(* IEC 61131-3 sources: plc-iiot-stack/src/POUs/Iiot/FB_MqttDiag, 14 files *)

(* ---- FB_MqttDiag.decl.st ---- *)
// Назначение: ведение связи с брокером и состояние узла (data_schema 6): автомат Disabled -> Connecting ->
//             Connected -> Backoff -> Connecting; тайм-аут подключения, пауза между попытками удваивается от
//             tBackoffMin до tBackoffMax и снова минимальна после tStable устойчивой связи. Перед Connect —
//             завещание (LWT) в <prefix>/<sNode>/status/connection: offline/lwt со временем подключения;
//             после подключения — рождение online/birth (source, sw_version, period_ms), затем xReady.
//             Выключение при связи — offline/shutdown, разрыв в следующем вызове. Без часов ПЛК обмен не
//             начинается (MQTT_ERR_NO_CLOCK). Счётчики, код последней ошибки, сводный статус в духе NE 107.
// Автор:      kr0nsch
// Версия:     0.1.0
// Документ:   docs/plc_mqtt.md, раздел «Связь и состояние узла»
FUNCTION_BLOCK FB_MqttDiag
VAR_INPUT
    xEnable : BOOL;
    itfClient : I_MqttClient;
    ltNow : LTIME;                                            // монотонное время (LTIME())
    uliTs_ms : ULINT;                                         // время UTC, мс (поле ts)
    sTopicPrefix : STRING(GVL_Const.IIOT_PREFIX_LEN);         // site/area/unit
    sNode : STRING(GVL_Const.IIOT_DEVICE_LEN) := 'PLC1';
    sSwVersion : STRING(GVL_Const.IIOT_TEXT_LEN) := '0.1.0';
    tPeriod : TIME := GVL_Const.TELEMETRY_PERIOD_DEFAULT;    // период контрольной публикации (period_ms)
    tConnectTimeout : TIME := GVL_Const.CONNECT_TIMEOUT_DEFAULT;
    tBackoffMin : TIME := GVL_Const.BACKOFF_MIN_DEFAULT;
    tBackoffMax : TIME := GVL_Const.BACKOFF_MAX_DEFAULT;
    tStable : TIME := GVL_Const.STABLE_TIME_DEFAULT;
    tDegradeWindow : TIME := GVL_Const.TELEMETRY_PERIOD_DEFAULT;   // окно оценки отказов публикаций
    uiFailThreshold : UINT := GVL_Const.FAIL_THRESHOLD_DEFAULT;
    udiPubFailed : UDINT;                                     // отказы публикаций телеметрии и тревог
END_VAR
VAR_IN_OUT
    stBroker : ST_MqttBrokerCfg;                              // ФБ дописывает топик и текст LWT
END_VAR
VAR_OUTPUT
    eState : E_MqttConnState := E_MqttConnState.Disabled;
    eNe107 : E_IiotNe107 := E_IiotNe107.CheckFunction;
    xConnected : BOOL;
    xReady : BOOL;                  // связь есть и рождение опубликовано: можно публиковать
    udiConnects : UDINT;            // успешных подключений
    udiDisconnects : UDINT;         // потерь установленной связи
    udiConnectFailures : UDINT;     // неудачных попыток подключения
    uiConsecutiveFailures : UINT;   // неудачных попыток подряд (сброс после tStable связи)
    diLastError : DINT;             // GVL_Const.MQTT_ERR_* или код библиотеки
    tBackoff : TIME;                // пауза перед следующей попыткой
    xDegraded : BOOL;               // за последнее окно публикации отклонялись
END_VAR
VAR
    ltStateSince : LTIME;
    ltDegradeStart : LTIME;
    udiPubFailedRef : UDINT;
    fbJson : FB_JsonBuilder;
    sTopic : STRING(GVL_Const.MQTT_TOPIC_LEN);
END_VAR

(* ---- BuildStatus.method.decl.st ---- *)
// JSON состояния узла в fbJson: online/birth (с source, sw_version, period_ms) или offline/<sReason>.
METHOD PRIVATE BuildStatus : BOOL
VAR_INPUT
    xOnline : BOOL;
    sReason : STRING(GVL_Const.IIOT_TEXT_LEN);
END_VAR

(* ---- BuildStatus.method.impl.st ---- *)
fbJson.Begin();
fbJson.AddString(sKey := 'schema_version', sValue := GVL_Const.IIOT_SCHEMA_VERSION);
fbJson.AddInt(sKey := 'ts', liValue := ULINT_TO_LINT(uliTs_ms));
fbJson.AddString(sKey := 'node', sValue := sNode);
IF xOnline THEN
    fbJson.AddString(sKey := 'state', sValue := 'online');
ELSE
    fbJson.AddString(sKey := 'state', sValue := 'offline');
END_IF
fbJson.AddString(sKey := 'reason', sValue := sReason);
IF xOnline THEN
    fbJson.AddString(sKey := 'source', sValue := GVL_Const.IIOT_SOURCE);
    fbJson.AddString(sKey := 'sw_version', sValue := sSwVersion);
    fbJson.AddInt(sKey := 'period_ms', liValue := ULINT_TO_LINT(TIME_TO_ULINT(tPeriod)));
END_IF
BuildStatus := fbJson.Finish();

(* ---- ConnectFailed.method.decl.st ---- *)
// Неудачная попытка подключения: код ошибки (клиента или diDefaultError), счётчики, разрыв, пауза.
METHOD PRIVATE ConnectFailed
VAR_INPUT
    diDefaultError : DINT;
END_VAR

(* ---- ConnectFailed.method.impl.st ---- *)
diLastError := itfClient.LastError();
IF diLastError = GVL_Const.MQTT_ERR_NONE THEN
    diLastError := diDefaultError;
END_IF
udiConnectFailures := udiConnectFailures + 1;
IF uiConsecutiveFailures < UINT#65535 THEN
    uiConsecutiveFailures := uiConsecutiveFailures + 1;
END_IF
itfClient.Disconnect();
EnterState(eNewState := E_MqttConnState.Backoff);

(* ---- EnterState.method.decl.st ---- *)
// Перейти в состояние eNewState и запомнить время входа.
METHOD PRIVATE EnterState
VAR_INPUT
    eNewState : E_MqttConnState;
END_VAR

(* ---- EnterState.method.impl.st ---- *)
IF eState <> eNewState THEN
    eState := eNewState;
    ltStateSince := ltNow;
END_IF

(* ---- FB_MqttDiag.impl.st ---- *)
// Выключено или нет часов: штатно закрыть связь (offline/shutdown, разрыв в следующем вызове)
IF NOT xEnable OR itfClient = 0 OR NOT F_IiotClockValid(uliTs_ms := uliTs_ms) THEN
    IF itfClient = 0 THEN
        EnterState(eNewState := E_MqttConnState.Disabled);
    ELSIF eState = E_MqttConnState.Connected AND xReady AND_THEN itfClient.IsConnected() THEN
        PublishStatus(xOnline := FALSE, sReason := 'shutdown');
        EnterState(eNewState := E_MqttConnState.Closing);
    ELSIF eState <> E_MqttConnState.Disabled THEN
        itfClient.Disconnect();
        EnterState(eNewState := E_MqttConnState.Disabled);
    END_IF
    IF xEnable AND NOT F_IiotClockValid(uliTs_ms := uliTs_ms) THEN
        diLastError := GVL_Const.MQTT_ERR_NO_CLOCK;
    END_IF
    uiConsecutiveFailures := 0;
    tBackoff := tBackoffMin;
    xConnected := FALSE;
    xReady := FALSE;
    xDegraded := FALSE;
    eNe107 := E_IiotNe107.CheckFunction;
    RETURN;
END_IF
IF tBackoff < tBackoffMin THEN
    tBackoff := tBackoffMin;
END_IF

CASE eState OF
    E_MqttConnState.Disabled, E_MqttConnState.Closing:
        IF eState = E_MqttConnState.Closing THEN
            itfClient.Disconnect();
        END_IF
        StartConnect(stBrokerCfg := stBroker);

    E_MqttConnState.Connecting:
        IF NOT itfClient.IsConnected() AND_THEN InState() >= TIME_TO_LTIME(tConnectTimeout) THEN
            ConnectFailed(diDefaultError := GVL_Const.MQTT_ERR_CONNECT_TIMEOUT);
        END_IF

    E_MqttConnState.Connected:
        IF NOT itfClient.IsConnected() THEN
            udiDisconnects := udiDisconnects + 1;
            diLastError := itfClient.LastError();
            IF diLastError = GVL_Const.MQTT_ERR_NONE THEN
                diLastError := GVL_Const.MQTT_ERR_CONNECTION_LOST;
            END_IF
            itfClient.Disconnect();
            xReady := FALSE;
            EnterState(eNewState := E_MqttConnState.Backoff);
        ELSIF InState() >= TIME_TO_LTIME(tStable) THEN
            // связь устойчива: следующая потеря — с минимальной паузы
            tBackoff := tBackoffMin;
            uiConsecutiveFailures := 0;
        END_IF

    E_MqttConnState.Backoff:
        IF InState() >= TIME_TO_LTIME(tBackoff) THEN
            // пауза для следующей неудачи — вдвое больше, не больше tBackoffMax
            IF tBackoff >= tBackoffMax / 2 THEN
                tBackoff := tBackoffMax;
            ELSE
                tBackoff := tBackoff * 2;
            END_IF
            StartConnect(stBrokerCfg := stBroker);
        END_IF
END_CASE

// подключение могло состояться в этом же вызове
IF eState = E_MqttConnState.Connecting AND_THEN itfClient.IsConnected() THEN
    udiConnects := udiConnects + 1;
    EnterState(eNewState := E_MqttConnState.Connected);
    xReady := FALSE;
    xDegraded := FALSE;
    ltDegradeStart := ltNow;
    udiPubFailedRef := udiPubFailed;
END_IF
xConnected := eState = E_MqttConnState.Connected;

// рождение узла, затем можно публиковать
IF xConnected AND NOT xReady THEN
    xReady := PublishStatus(xOnline := TRUE, sReason := 'birth');
END_IF
// отказы публикаций за окно
IF xConnected THEN
    IF ltNow < ltDegradeStart THEN
        ltDegradeStart := ltNow;
    ELSIF (ltNow - ltDegradeStart) >= TIME_TO_LTIME(tDegradeWindow) THEN
        ltDegradeStart := ltNow;
        xDegraded := udiPubFailed <> udiPubFailedRef;
        udiPubFailedRef := udiPubFailed;
    END_IF
END_IF
UpdateNe107();

(* ---- InState.method.impl.st ---- *)
IF ltNow < ltStateSince THEN
    ltStateSince := ltNow;
END_IF
InState := ltNow - ltStateSince;

(* ---- PublishStatus.method.decl.st ---- *)
// Опубликовать состояние узла (QoS 1, retain). TRUE — клиент принял.
METHOD PRIVATE PublishStatus : BOOL
VAR_INPUT
    xOnline : BOOL;
    sReason : STRING(GVL_Const.IIOT_TEXT_LEN);
END_VAR

(* ---- PublishStatus.method.impl.st ---- *)
sTopic := StatusTopic();
IF NOT BuildStatus(xOnline := xOnline, sReason := sReason) OR LEN(sTopic) = 0 THEN
    RETURN;
END_IF
PublishStatus := itfClient.Publish(sTopic := sTopic, eQos := E_MqttQos.AtLeastOnce, xRetain := TRUE,
                                   sPayload := fbJson.sJson);

(* ---- StartConnect.method.decl.st ---- *)
// Завещание offline/lwt со временем подключения в параметрах брокера и запрос подключения; отказ клиента —
// неудачная попытка.
METHOD PRIVATE StartConnect
VAR_IN_OUT
    stBrokerCfg : ST_MqttBrokerCfg;
END_VAR

(* ---- StartConnect.method.impl.st ---- *)
stBrokerCfg.sWillTopic := StatusTopic();
IF BuildStatus(xOnline := FALSE, sReason := 'lwt') THEN
    stBrokerCfg.sWillPayload := fbJson.sJson;
ELSE
    stBrokerCfg.sWillPayload := '';
END_IF
stBrokerCfg.xWillRetain := TRUE;
EnterState(eNewState := E_MqttConnState.Connecting);
IF NOT itfClient.Connect(stCfg := stBrokerCfg) THEN
    ConnectFailed(diDefaultError := GVL_Const.MQTT_ERR_CONNECT_REJECTED);
END_IF

(* ---- UpdateNe107.method.impl.st ---- *)
CASE eState OF
    E_MqttConnState.Disabled, E_MqttConnState.Closing:
        eNe107 := E_IiotNe107.CheckFunction;
    E_MqttConnState.Connected:
        IF xDegraded THEN
            eNe107 := E_IiotNe107.MaintenanceRequired;
        ELSE
            eNe107 := E_IiotNe107.Good;
        END_IF
ELSE
    IF uiConsecutiveFailures >= MAX(uiFailThreshold, 1) THEN
        eNe107 := E_IiotNe107.Failure;
    ELSIF udiConnects = 0 AND uiConsecutiveFailures = 0 THEN
        eNe107 := E_IiotNe107.CheckFunction;
    ELSE
        eNe107 := E_IiotNe107.OutOfSpecification;
    END_IF
END_CASE
